FUNCTION_BLOCK FB_RelayBistableToggle IMPLEMENTS I_Relay
VAR_INPUT
    stDeviceId : ST_DeviceId;
END_VAR
VAR_OUTPUT
    bTogglePulse : BOOL;
END_VAR
VAR
    bRequestedState : BOOL;
    bCurrentState   : BOOL;
    fbTrigger       : R_TRIG;
    fbPulse         : TP;
END_VAR

fbTrigger(CLK := (bRequestedState <> bCurrentState) AND NOT fbPulse.Q);
fbPulse(IN := fbTrigger.Q, PT := T#100MS);

IF fbTrigger.Q THEN
    bCurrentState := bRequestedState;
END_IF

bTogglePulse := fbPulse.Q;

PROPERTY DeviceId : ST_DeviceId
GET
DeviceId := stDeviceId;
END_GET
END_PROPERTY

PROPERTY IsOn : BOOL
GET
IsOn := bCurrentState;
END_GET
END_PROPERTY

METHOD PUBLIC TurnOn
bRequestedState := TRUE;
END_METHOD

METHOD PUBLIC TurnOff
bRequestedState := FALSE;
END_METHOD

METHOD PUBLIC Toggle
bRequestedState := NOT bRequestedState;
END_METHOD

END_FUNCTION_BLOCK

(* stored: Version 1.1.0.1, ProductVersion 3.1.4026.20
   POU FB_RelayBistableToggle: Id {88888888-8888-4888-8888-888888888880}
   Property DeviceId: Id {88888888-0000-4000-8000-000000000001}
   Get Get: Id {88888888-0000-4000-8000-000000000011}
   Property IsOn: Id {88888888-0000-4000-8000-000000000002}
   Get Get: Id {88888888-0000-4000-8000-000000000012}
   Method TurnOn: Id {88888888-0000-4000-8000-000000000003}
   Method TurnOff: Id {88888888-0000-4000-8000-000000000004}
   Method Toggle: Id {88888888-0000-4000-8000-000000000005} *)
